Fanuc KAREL source: KT00817.KL

PROGRAM KT00817
%NOLOCKGROUP
VAR
  B1: BOOLEAN
  B2: BOOLEAN
  OUT: REAL
BEGIN
  B1 = TRUE
  B2 = FALSE
  B1 = TRUE
  B2 = FALSE
  OUT = LN(B1)
END KT00817
